(*
SPDX-FileCopyrightText: © 2026 Oleksandr Tiutyk <trofimich@gmail.com>
SPDX-License-Identifier: MIT
License: https://opensource.org/license/mit
*)

(*!
<summary>Shows a complete single-cycle test body without guards or contexts.</summary>
*)

{attribute 'no_explicit_call' := 'do not call this function block directly'}
FUNCTION_BLOCK AdditionTest EXTENDS TOF_Testing.SingleCycleTest
VAR_STAT
	{attribute 'hide'}
	_ClassName : STRING := __POUNAME();
END_VAR

//! <summary>Borrows the concrete class name for the lifetime of this instance; callers must not modify it.</summary>
{attribute 'monitoring' := 'call'}
PROPERTY ClassName : REFERENCE TO STRING
GET
ClassName REF= _ClassName;
END_GET
END_PROPERTY

(*!
<summary>Checks an arithmetic result and completes automatically on return.</summary>
*)
METHOD PROTECTED ExecuteTest
Assert.ThatDInt(actual := 2 + 3).ToBe(expected := 5);
END_METHOD

//! <summary>Borrows the compiler-initialized namespace; callers must not modify the returned reference.</summary>
{attribute 'monitoring' := 'call'}
PROPERTY NamespaceName : REFERENCE TO STRING
GET
NamespaceName REF= CurrentNamespace.Name;
END_GET
END_PROPERTY

//! <summary>Reports the complete concrete instance size, excluding separately allocated storage.</summary>
{attribute 'monitoring' := 'call'}
PROPERTY SelfSize : ULINT
GET
SelfSize := XSIZEOF(THIS^);
END_GET
END_PROPERTY

END_FUNCTION_BLOCK

(* stored: Version 1.1.0.1
   POU AdditionTest: Id {8be6ae55-55a0-4318-ac83-0314063ff386}, SpecialFunc None
   Property ClassName: Id {d4e36c71-455c-41e8-90bc-3b278a4769d4}
   Get Get: Id {4396c153-2d9a-44a3-b477-9a38834b2bf4}
   Method ExecuteTest: Id {bed355e0-44ef-4446-9d12-1a3dbd028abc}
   Property NamespaceName: Id {dcce0949-f2cb-4d4a-ad0c-b60bcc319dba}
   Get Get: Id {3bdae836-0be2-4f4f-90a7-574ca91995de}
   Property SelfSize: Id {5413998b-7a75-4baa-a6d3-0ed4dd5fd06b}
   Get Get: Id {8dc944d1-fccb-49f9-9046-3c8a06dec385} *)
